Fanuc KAREL source: KT00570.KL

PROGRAM KT00570
%NOLOCKGROUP
VAR
  V1: VECTOR
  R2: REAL
  OUT: VECTOR
BEGIN
  V1.X = 1.0
    R2 = 3.0
  OUT = V1 @ R2
END KT00570
